// Common part of catalog alarms and messages.
INTERFACE I_CatalogEvent

PROPERTY Arguments : I_ArgumentBuilder
GET
END_GET
END_PROPERTY

PROPERTY Severity : TcEventSeverity
GET
END_GET
END_PROPERTY

PROPERTY LastResult : HRESULT
GET
END_GET
END_PROPERTY

PROPERTY SourceName : T_MaxString
GET
END_GET
SET
END_SET
END_PROPERTY

END_INTERFACE

(* stored: Version 1.1.0.1, ProductVersion 3.1.4026.26
   Itf I_CatalogEvent: Id {ecbf0128-e578-407b-9065-9e0b8dda54a4}
   Property Arguments: Id {dfac73f4-e1e7-4f41-bea0-76fb726d7ee9}
   Get Get: Id {1d362b96-2755-44c5-af99-faa5daa4ee0e}
   Property Severity: Id {79a4b9a6-24e2-42c9-8f58-59cebe64b57d}
   Get Get: Id {c28f00d7-06a8-4080-b533-d2f64f2bc7b6}
   Property LastResult: Id {8a16e2e3-0488-4c34-81a4-8fdefc5af7ac}
   Get Get: Id {65dd371c-a6ca-4be0-92fa-11b77ba3a6ea}
   Property SourceName: Id {c8a97ec5-4e4d-42df-a292-6bbde6abcf9b}
   Get Get: Id {86395133-2cd1-4f65-b3c7-4efa6a54af9d}
   Set Set: Id {1958da8b-7472-4cad-9714-7c8905e0612a} *)
